TYPE "UDT_Service_ValueDefinition"
VERSION : 0.1
   STRUCT
      indexMTP : Int;   // MTP Index of value
      indexIO : Int;   // IO Index of value
      "type" : Int;   // Type of parameter
      controlModule : Byte := 16#FF;   // Number of control module used with parameter
   END_STRUCT;

END_TYPE

